Fanuc KAREL source: KT00227.KL

PROGRAM KT00227
%NOLOCKGROUP
VAR
  B1: BOOLEAN
  I2: INTEGER
  OUT: BOOLEAN
BEGIN
  B1 = TRUE
    I2 = 3
  OUT = B1 OR I2
END KT00227
